(* IEC 61131-3 sources: llm-plc-st-eval/data/processed_v2_primera/claude-sonnet-4-6/B3/zero_shot, 3 files *)

(* ---- ejec_1.st ---- *)
FUNCTION_BLOCK FB_Contador
VAR_INPUT
    sensorPieza : BOOL; (* Señal del sensor fotoeléctrico *)
    btnReset    : BOOL; (* Botón de reset de la cuenta *)
END_VAR

VAR_OUTPUT
    loteListo : BOOL; (* Activa cuando se completan 12 piezas *)
    cuenta    : INT;  (* Número de piezas contadas *)
END_VAR

VAR
    sensorPiezaPrev : BOOL; (* Estado anterior del sensor para detección de flanco *)
END_VAR

(* ─────────────────────────────────────────────
   Constantes
   ───────────────────────────────────────────── *)
VAR CONSTANT
    TAMANO_LOTE : INT := 12; (* Piezas por lote *)
END_VAR

(* ══════════════════════════════════════════════
   LÓGICA PRINCIPAL
   ══════════════════════════════════════════════ *)

(* 1. Reset: tiene prioridad sobre el conteo *)
IF btnReset THEN
    cuenta        := 0;
    loteListo     := FALSE;
    sensorPiezaPrev := FALSE;

(* 2. Conteo normal: solo si el lote no está completo *)
ELSIF NOT loteListo THEN

    (* Detectar flanco ascendente del sensor (FALSE → TRUE) *)
    IF sensorPieza AND NOT sensorPiezaPrev THEN
        cuenta := cuenta + 1;
    END_IF;

    (* Activar salida cuando se alcanza el tamaño de lote *)
    IF cuenta >= TAMANO_LOTE THEN
        loteListo := TRUE;
    END_IF;

END_IF;

(* 3. Guardar estado actual del sensor para el próximo ciclo *)
sensorPiezaPrev := sensorPieza;

(* ---- ejec_2.st ---- *)
FUNCTION_BLOCK FB_Contador
VAR_INPUT
    sensorPieza : BOOL; (* Señal del sensor fotoeléctrico *)
    btnReset    : BOOL; (* Botón de reset de cuenta y lote *)
END_VAR

VAR_OUTPUT
    loteListo : BOOL; (* Activa cuando se completan 12 piezas *)
    cuenta    : INT;  (* Número de piezas contadas *)
END_VAR

VAR
    sensorPiezaAnterior : BOOL; (* Valor previo del sensor para detectar flanco *)
END_VAR

(* ── Constantes ── *)
VAR CONSTANT
    TAMANO_LOTE : INT := 12; (* Número de piezas por lote *)
END_VAR

(* ════════════════════════════════════════════════════════
   Lógica principal
   ════════════════════════════════════════════════════════ *)

(* 1. Reset: prioridad alta sobre el conteo *)
IF btnReset THEN
    cuenta    := 0;
    loteListo := FALSE;

ELSE
    (* 2. Detección de flanco ascendente del sensor (FALSE → TRUE) *)
    IF sensorPieza AND NOT sensorPiezaAnterior THEN
        (* Solo contar si el lote aún no está completo *)
        IF NOT loteListo THEN
            cuenta := cuenta + 1;
        END_IF;
    END_IF;

    (* 3. Activar salida de lote al alcanzar el tamaño definido *)
    IF cuenta >= TAMANO_LOTE THEN
        loteListo := TRUE;
    END_IF;
END_IF;

(* 4. Actualizar memoria de flanco para el próximo ciclo *)
sensorPiezaAnterior := sensorPieza;

(* ---- ejec_3.st ---- *)
FUNCTION_BLOCK FB_Contador
VAR_INPUT
    sensorPieza : BOOL; (* Señal del sensor fotoeléctrico *)
    btnReset    : BOOL; (* Botón de reset de la cuenta *)
END_VAR

VAR_OUTPUT
    loteListo : BOOL; (* TRUE cuando se completan 12 piezas *)
    cuenta    : INT;  (* Contador de piezas detectadas *)
END_VAR

VAR
    sensorPiezaPrev : BOOL; (* Estado anterior del sensor para detección de flanco *)
END_VAR

(* ─────────────────────────────────────────────
   Constantes de configuración
   ───────────────────────────────────────────── *)
VAR CONSTANT
    TAMANO_LOTE : INT := 12; (* Número de piezas por lote *)
END_VAR

(* ══════════════════════════════════════════════
   LÓGICA PRINCIPAL
   ══════════════════════════════════════════════ *)

(* 1. Reset: tiene prioridad sobre el conteo *)
IF btnReset THEN
    cuenta         := 0;
    loteListo      := FALSE;
    sensorPiezaPrev := FALSE;

(* 2. Conteo activo solo si el lote no está completo *)
ELSIF NOT loteListo THEN

    (* Detección de flanco ascendente del sensor (FALSE → TRUE) *)
    IF sensorPieza AND NOT sensorPiezaPrev THEN
        cuenta := cuenta + 1;
    END_IF;

    (* Activar salida cuando se alcanza el tamaño de lote *)
    IF cuenta >= TAMANO_LOTE THEN
        loteListo := TRUE;
    END_IF;

END_IF;

(* 3. Actualizar estado previo del sensor *)
sensorPiezaPrev := sensorPieza;
